(*
SPDX-FileCopyrightText: © 2026 Oleksandr Tiutyk <trofimich@gmail.com>
SPDX-License-Identifier: MIT
License: https://opensource.org/license/mit
*)

(*!
<summary>Observes workflow hooks and injects one recoverable initialization failure.</summary>
<description>
Variable storage belongs to this persistent fixture. The initialization failure is raised only after one
ordinary binding was added, allowing the caller to observe the configured retry policy.
</description>
*)

{attribute 'no_explicit_call' := 'do not call this function block directly'}
{attribute 'no_assign'}
FUNCTION_BLOCK WorkflowContractWorkflow EXTENDS TOF_Workflow.Workflow
VAR_INPUT
	//! <summary>Raises once after registering the initialization binding.</summary>
	throwInitialization : BOOL;
END_VAR
VAR_OUTPUT
	//! <summary>Total calls to InitializeVariables.</summary>
	initializationCount : DINT;
	//! <summary>Total calls to OnAfterRootActivityExecute.</summary>
	afterCount : DINT;
END_VAR
VAR_STAT
	//! <summary>Distinct static field to avoid redeclaring inherited Workflow metadata.</summary>
	_ProbeClassName : STRING := __POUNAME();
END_VAR
VAR
	_RegisteredValue : DINT;
END_VAR

(*!
<summary>Returns the initialized static name of this concrete fixture.</summary>
*)
{attribute 'monitoring' := 'call'}
PROPERTY ClassName : REFERENCE TO STRING
GET
ClassName REF= _ProbeClassName;
END_GET
END_PROPERTY

(*!
<summary>Borrows the test project namespace without changing it.</summary>
*)
{attribute 'monitoring' := 'call'}
PROPERTY NamespaceName : REFERENCE TO STRING
GET
// SA0006: Read-only namespace string borrowed across test tasks.
{analysis -6}
NamespaceName REF= CurrentNamespace.Name;
{analysis +6}
END_GET
END_PROPERTY

(*!
<summary>Reports the size of this concrete fixture in bytes.</summary>
*)
{attribute 'monitoring' := 'call'}
PROPERTY SelfSize : ULINT
GET
SelfSize := XSIZEOF(THIS^);
END_GET
END_PROPERTY

(*!
<summary>Registers persistent fixture storage and optionally interrupts the first attempt.</summary>
*)
METHOD PROTECTED InitializeVariables
initializationCount := initializationCount + 1;
BindPlcVariable(name := 'Initialized', plcVariable := _RegisteredValue);

IF throwInitialization THEN
	throwInitialization := FALSE;

	TOF_Core.Exceptions.ThrowStandard(
		sourceNamespaceName := NamespaceName,
		sourceClassName := ClassName,
		sourcePOUName := __POUNAME(),
		sourcePosition := __POSITION(),
		message := "Controlled variable initialization failure"
	);
END_IF
END_METHOD

(*!
<summary>Counts completion of the workflow execution boundary.</summary>
*)
METHOD PROTECTED OnAfterRootActivityExecute
afterCount := afterCount + 1;
END_METHOD

END_FUNCTION_BLOCK

(* stored: Version 1.1.0.1
   POU WorkflowContractWorkflow: Id {b6ce7c43-77ab-4ec3-b8f2-3fabd09b4738}, SpecialFunc None
   Property ClassName: Id {f1c20fed-4365-4054-bfed-dd49b242f3b5}
   Get Get: Id {02181012-bc3e-447a-a7c4-b88cde090f5c}
   Property NamespaceName: Id {b36792f7-f1bd-4687-b0d7-a3a701165a55}
   Get Get: Id {26d36206-9d76-4ab1-8d37-92b65a0a404c}
   Property SelfSize: Id {9d992b5a-e449-4301-904d-dbe8afb5952e}
   Get Get: Id {f4e8703b-6af3-4cf4-a847-7bf995e49da1}
   Method InitializeVariables: Id {ffd75302-3b07-47f3-ad22-b2413fe6b079}
   Method OnAfterRootActivityExecute: Id {445fe8bb-c2a7-4429-9199-4a91e3760d3f} *)
